Fanuc KAREL source: KO00107.KL

PROGRAM KO00107
%NOLOCKGROUP
VAR
  A: REAL
  B: REAL
  OUT: INTEGER
BEGIN
  A = 1
  B = 2
  OUT = ATAN2(A, B)
END KO00107
